(* IEC 61131-3 sources: codesys-framework/txt/application/WeVe General (library)/Blink/DUT, 1 file *)

(* ---- SC_Blinks.dut.st ---- *)
TYPE SC_Blinks :
STRUCT

	xBlink200msLow1800msHigh 		: BOOL;
	xBlink1800msLow200msHigh 		: BOOL;
	xBlink1000msLow1000msHigh 		: BOOL;
	xBlink250msLow250msHigh 		: BOOL;
	xBlink500msLow500msHigh 		: BOOL;
	xBlink100msLow100msHigh 		: BOOL;

END_STRUCT
END_TYPE
